(****************************************************************************************************<br>
© Syntegon Group.<br>
All rights reserved, also regarding any disposal, exploitation, reproduction, editing, distribution,<br>
as well as in the event of applications for industrial property rights.<br>
*****************************************************************************************************<br>
DESCRIPTION:<br>
Base of every robot (Delta, XTS gantry, XTS loop, Cartesian): zones plus the gripper fingers, m_SetFinger,<br>
m_SetFingerOffset (a finger's place on the flange) and m_ClearFingers, the limit area, m_SetLimitArea and<br>
m_ClearLimitArea, and the TCP limit area, m_SetTcpLimitArea and m_ClearTcpLimitArea. A derived FB tells where<br>
its fingers and its boxes lie through m_Fingers and m_LimitArea; an XTS loop has neither box.<br>
Not used directly.<br>
*****************************************************************************************************<br>
VERSION         ¦ DATE       ¦ NAME      ¦ CHANGE<br>
Syn_Visu 4.0.0  ¦ 2026-11-01 ¦ J.Willner ¦ New: fingers shared by all robots<br>
Syn_Visu 9.3.0  ¦ 2026-11-07 ¦ J.Willner ¦ Limit area shared by Delta, XTS gantry and Cartesian (was Delta only)<br>
Syn_Visu 9.4.0  ¦ 2026-11-09 ¦ J.Willner ¦ TCP limit area: m_SetTcpLimitArea, m_ClearTcpLimitArea<br>
Syn_Visu 9.4.1  ¦ 2026-11-09 ¦ J.Willner ¦ Limit area compares ignore padding: no config change from unchanged values<br>
Syn_Visu 9.5.0  ¦ 2026-11-11 ¦ J.Willner ¦ m_SetFingerOffset: a finger's place on the flange (ADR 0018)<br>
****************************************************************************************************)
FUNCTION_BLOCK ABSTRACT _FB_VisuRobot EXTENDS _FB_VisuZoneComponent

(****************************************************************************************************<br>
© Syntegon Group.<br>
All rights reserved, also regarding any disposal, exploitation, reproduction, editing, distribution,<br>
as well as in the event of applications for industrial property rights.<br>
*****************************************************************************************************<br>
DESCRIPTION:<br>
Removes the gripper definition. TRUE if there was one.<br>
****************************************************************************************************)
METHOD m_ClearFingers : BOOL
VAR
	p_TempCount							: POINTER TO UINT;
	p_TempFingers						: POINTER TO ARRAY[0..VISU_GlobalConst_Param.VISU_un_MAX_FINGERS - 1] OF ST_VisuFinger;
	TempEmpty							: ST_VisuFinger;
	un_TempIndex						: UINT;
END_VAR
m_ClearFingers := FALSE;
m_Fingers(vo_p_Count => p_TempCount, vo_p_Fingers => p_TempFingers);
IF p_TempCount = 0 OR p_TempFingers = 0 THEN
	RETURN;
END_IF
m_ClearFingers := p_TempCount^ > 0;
FOR un_TempIndex := 0 TO VISU_GlobalConst_Param.VISU_un_MAX_FINGERS - 1 DO
	p_TempFingers^[un_TempIndex] := TempEmpty;
END_FOR
p_TempCount^ := 0;
IF m_ClearFingers THEN
	m_NotifyConfigChanged();
END_IF
END_METHOD

(****************************************************************************************************<br>
© Syntegon Group.<br>
All rights reserved, also regarding any disposal, exploitation, reproduction, editing, distribution,<br>
as well as in the event of applications for industrial property rights.<br>
*****************************************************************************************************<br>
DESCRIPTION:<br>
Removes the limit area. TRUE if there was one.<br>
****************************************************************************************************)
METHOD m_ClearLimitArea : BOOL
VAR
	p_TempLimitArea						: POINTER TO ST_VisuLimitArea;
	TempEmpty							: ST_VisuLimitArea;
END_VAR
m_ClearLimitArea := FALSE;
m_LimitArea(vo_p_LimitArea => p_TempLimitArea);
IF p_TempLimitArea = 0 THEN
	RETURN;
END_IF
m_ClearLimitArea := p_TempLimitArea^.bActive;
(* Zeroed first: the MEMCMP below also compares the padding after bActive, which a method local leaves undefined. *)
Tc2_System.MEMSET(ADR(TempEmpty), 0, SIZEOF(TempEmpty));
IF Tc2_System.MEMCMP(ADR(TempEmpty), p_TempLimitArea, SIZEOF(TempEmpty)) <> 0 THEN
	p_TempLimitArea^ := TempEmpty;
	m_NotifyConfigChanged();
END_IF
END_METHOD

(****************************************************************************************************<br>
© Syntegon Group.<br>
All rights reserved, also regarding any disposal, exploitation, reproduction, editing, distribution,<br>
as well as in the event of applications for industrial property rights.<br>
*****************************************************************************************************<br>
DESCRIPTION:<br>
Removes the TCP limit area. TRUE if there was one.<br>
****************************************************************************************************)
METHOD m_ClearTcpLimitArea : BOOL
VAR
	p_TempTcpLimitArea					: POINTER TO ST_VisuLimitArea;
	TempEmpty							: ST_VisuLimitArea;
END_VAR
m_ClearTcpLimitArea := FALSE;
m_LimitArea(vo_p_TcpLimitArea => p_TempTcpLimitArea);
IF p_TempTcpLimitArea = 0 THEN
	RETURN;
END_IF
m_ClearTcpLimitArea := p_TempTcpLimitArea^.bActive;
(* Zeroed first: the MEMCMP below also compares the padding after bActive, which a method local leaves undefined. *)
Tc2_System.MEMSET(ADR(TempEmpty), 0, SIZEOF(TempEmpty));
IF Tc2_System.MEMCMP(ADR(TempEmpty), p_TempTcpLimitArea, SIZEOF(TempEmpty)) <> 0 THEN
	p_TempTcpLimitArea^ := TempEmpty;
	m_NotifyConfigChanged();
END_IF
END_METHOD

(****************************************************************************************************<br>
© Syntegon Group.<br>
All rights reserved, also regarding any disposal, exploitation, reproduction, editing, distribution,<br>
as well as in the event of applications for industrial property rights.<br>
*****************************************************************************************************<br>
DESCRIPTION:<br>
Where the gripper fingers lie in the derived FB's contract structure: vo_p_Count points to its<br>
nFingerCount, vo_p_Fingers to its aFingers.<br>
****************************************************************************************************)
METHOD PROTECTED ABSTRACT m_Fingers : BOOL
VAR_OUTPUT
	vo_p_Count							: POINTER TO UINT;
	vo_p_Fingers						: POINTER TO ARRAY[0..VISU_GlobalConst_Param.VISU_un_MAX_FINGERS - 1] OF ST_VisuFinger;
END_VAR
END_METHOD

(****************************************************************************************************<br>
© Syntegon Group.<br>
All rights reserved, also regarding any disposal, exploitation, reproduction, editing, distribution,<br>
as well as in the event of applications for industrial property rights.<br>
*****************************************************************************************************<br>
DESCRIPTION:<br>
Where the limit area and the TCP limit area lie in the derived FB's contract structure: vo_p_LimitArea points<br>
to its stLimitArea, vo_p_TcpLimitArea to its stTcpLimitArea; both are 0 for a robot without them (XTS loop: it<br>
has no working area of its own).<br>
****************************************************************************************************)
METHOD PROTECTED ABSTRACT m_LimitArea : BOOL
VAR_OUTPUT
	vo_p_LimitArea						: POINTER TO ST_VisuLimitArea;
	vo_p_TcpLimitArea					: POINTER TO ST_VisuLimitArea;
END_VAR
END_METHOD

(****************************************************************************************************<br>
© Syntegon Group.<br>
All rights reserved, also regarding any disposal, exploitation, reproduction, editing, distribution,<br>
as well as in the event of applications for industrial property rights.<br>
*****************************************************************************************************<br>
DESCRIPTION:<br>
Defines gripper finger vi_un_Finger (1-based): a cylinder hanging from the finger's pose along its local -Z.<br>
For XTS kinematics it is a finger of every mover's gripper. The finger count grows to vi_un_Finger.<br>
Its place on the gripper flange comes from m_SetFingerOffset and is kept here.<br>
*****************************************************************************************************<br>
OUTPUT VALUES:<br>
FALSE outside 1..VISU_GlobalConst_Param.VISU_un_MAX_FINGERS.<br>
****************************************************************************************************)
METHOD m_SetFinger : BOOL
VAR_INPUT
	vi_un_Finger						: UINT;	// [-] 1-based, as a product's nFingerId
	vi_lr_Diameter						: LREAL;	// [mm]
	vi_lr_Height						: LREAL;	// [mm] along the finger's local -Z
END_VAR
VAR
	p_TempCount							: POINTER TO UINT;
	p_TempFingers						: POINTER TO ARRAY[0..VISU_GlobalConst_Param.VISU_un_MAX_FINGERS - 1] OF ST_VisuFinger;
	TempFinger							: ST_VisuFinger;
END_VAR
m_SetFinger := FALSE;
IF vi_un_Finger = 0 OR vi_un_Finger > VISU_GlobalConst_Param.VISU_un_MAX_FINGERS THEN
	RETURN;
END_IF
m_Fingers(vo_p_Count => p_TempCount, vo_p_Fingers => p_TempFingers);
IF p_TempCount = 0 OR p_TempFingers = 0 THEN
	RETURN;
END_IF
TempFinger.fDiameter := vi_lr_Diameter;
TempFinger.fHeight := vi_lr_Height;
(* The offset stays as m_SetFingerOffset set it. *)
TempFinger.stOffset := p_TempFingers^[vi_un_Finger - 1].stOffset;
IF vi_un_Finger > p_TempCount^
OR Tc2_System.MEMCMP(ADR(TempFinger), ADR(p_TempFingers^[vi_un_Finger - 1]), SIZEOF(TempFinger)) <> 0
THEN
	p_TempFingers^[vi_un_Finger - 1] := TempFinger;
	p_TempCount^ := MAX(p_TempCount^, vi_un_Finger);
	m_NotifyConfigChanged();
END_IF
m_SetFinger := TRUE;
END_METHOD

(****************************************************************************************************<br>
© Syntegon Group.<br>
All rights reserved, also regarding any disposal, exploitation, reproduction, editing, distribution,<br>
as well as in the event of applications for industrial property rights.<br>
*****************************************************************************************************<br>
DESCRIPTION:<br>
Places finger vi_un_Finger (1-based, defined with m_SetFinger) on the gripper flange (ADR 0018): the position<br>
of its frame in the flange frame and its rotation about the flange's Z. The flange frame's -Z points to the<br>
product: a Delta's lies at the TCP with the robot's axes, a Cartesian robot's has the robot's axes, an XTS mover's<br>
turns with the mover. While the application reports no pose for the finger (m_SetFingerState, or an XTS track<br>
with m_SetFingersOnFlange), the visualisation draws it there. The config version only changes when a value does.<br>
*****************************************************************************************************<br>
OUTPUT VALUES:<br>
FALSE for a finger outside 1..the finger count.<br>
****************************************************************************************************)
METHOD m_SetFingerOffset : BOOL
VAR_INPUT
	vi_un_Finger						: UINT;	// [-] 1-based
	vi_lr_X								: LREAL;	// [mm] along the flange's X
	vi_lr_Y								: LREAL;	// [mm] along the flange's Y
	vi_lr_Z								: LREAL;	// [mm] along the flange's Z (towards the product: negative)
	vi_lr_Rz							: LREAL;	// [deg] about the flange's Z
END_VAR
VAR
	p_TempCount							: POINTER TO UINT;
	p_TempFingers						: POINTER TO ARRAY[0..VISU_GlobalConst_Param.VISU_un_MAX_FINGERS - 1] OF ST_VisuFinger;
	TempOffset							: ST_VisuPlanarPose;
END_VAR
m_SetFingerOffset := FALSE;
m_Fingers(vo_p_Count => p_TempCount, vo_p_Fingers => p_TempFingers);
IF p_TempCount = 0 OR p_TempFingers = 0 THEN
	RETURN;
END_IF
IF vi_un_Finger = 0 OR vi_un_Finger > p_TempCount^ THEN
	RETURN;
END_IF
TempOffset.fX := vi_lr_X;
TempOffset.fY := vi_lr_Y;
TempOffset.fZ := vi_lr_Z;
TempOffset.fRz := vi_lr_Rz;
IF Tc2_System.MEMCMP(ADR(TempOffset), ADR(p_TempFingers^[vi_un_Finger - 1].stOffset), SIZEOF(TempOffset)) <> 0 THEN
	p_TempFingers^[vi_un_Finger - 1].stOffset := TempOffset;
	m_NotifyConfigChanged();
END_IF
m_SetFingerOffset := TRUE;
END_METHOD

(****************************************************************************************************<br>
© Syntegon Group.<br>
All rights reserved, also regarding any disposal, exploitation, reproduction, editing, distribution,<br>
as well as in the event of applications for industrial property rights.<br>
*****************************************************************************************************<br>
DESCRIPTION:<br>
Sets and activates the limit area: an axis-aligned box in the robot frame (relative to its pose, the frame its<br>
working area is given in) that further restricts the working area. Delta, XTS gantry and Cartesian robot;<br>
an XTS loop has none. Equal bounds make a flat box. The config version only changes when a value does.<br>
*****************************************************************************************************<br>
OUTPUT VALUES:<br>
TRUE if anything changed; FALSE for a robot without a limit area (XTS loop).<br>
****************************************************************************************************)
METHOD m_SetLimitArea : BOOL
VAR_INPUT
	vi_lr_XMin							: LREAL;	// [mm] in the robot frame
	vi_lr_XMax							: LREAL;	// [mm]
	vi_lr_YMin							: LREAL;	// [mm]
	vi_lr_YMax							: LREAL;	// [mm]
	vi_lr_ZMin							: LREAL;	// [mm] relative to the pose (below it: negative)
	vi_lr_ZMax							: LREAL;	// [mm]
END_VAR
VAR
	p_TempLimitArea						: POINTER TO ST_VisuLimitArea;
	TempLimitArea						: ST_VisuLimitArea;
END_VAR
m_SetLimitArea := FALSE;
m_LimitArea(vo_p_LimitArea => p_TempLimitArea);
IF p_TempLimitArea = 0 THEN
	RETURN;
END_IF
(* Zeroed first: the MEMCMP below also compares the padding after bActive, which a method local leaves undefined. *)
Tc2_System.MEMSET(ADR(TempLimitArea), 0, SIZEOF(TempLimitArea));
TempLimitArea.fXMin := vi_lr_XMin;
TempLimitArea.fXMax := vi_lr_XMax;
TempLimitArea.fYMin := vi_lr_YMin;
TempLimitArea.fYMax := vi_lr_YMax;
TempLimitArea.fZMin := vi_lr_ZMin;
TempLimitArea.fZMax := vi_lr_ZMax;
TempLimitArea.bActive := TRUE;
IF Tc2_System.MEMCMP(ADR(TempLimitArea), p_TempLimitArea, SIZEOF(TempLimitArea)) <> 0 THEN
	p_TempLimitArea^ := TempLimitArea;
	m_NotifyConfigChanged();
	m_SetLimitArea := TRUE;
END_IF
END_METHOD

(****************************************************************************************************<br>
© Syntegon Group.<br>
All rights reserved, also regarding any disposal, exploitation, reproduction, editing, distribution,<br>
as well as in the event of applications for industrial property rights.<br>
*****************************************************************************************************<br>
DESCRIPTION:<br>
Sets and activates the TCP limit area: an axis-aligned box around the TCP (XTS gantry: around every mover's<br>
gripper flange), its bounds relative to the TCP along the axes of the robot frame. It moves with the TCP and<br>
never turns. The visualisation lights it up red with a message when it overlaps another robot's limit area or<br>
TCP limit area (also another mover's of the same gantry), or leaves the robot's own limit area. Delta, XTS<br>
gantry and Cartesian robot; an XTS loop has none. Equal bounds make a flat box. The config version only<br>
changes when a value does.<br>
*****************************************************************************************************<br>
OUTPUT VALUES:<br>
TRUE if anything changed; FALSE for a robot without a TCP limit area (XTS loop).<br>
****************************************************************************************************)
METHOD m_SetTcpLimitArea : BOOL
VAR_INPUT
	vi_lr_XMin							: LREAL;	// [mm] relative to the TCP, along the robot frame's X
	vi_lr_XMax							: LREAL;	// [mm]
	vi_lr_YMin							: LREAL;	// [mm]
	vi_lr_YMax							: LREAL;	// [mm]
	vi_lr_ZMin							: LREAL;	// [mm] relative to the TCP (below it: negative)
	vi_lr_ZMax							: LREAL;	// [mm]
END_VAR
VAR
	p_TempTcpLimitArea					: POINTER TO ST_VisuLimitArea;
	TempTcpLimitArea					: ST_VisuLimitArea;
END_VAR
m_SetTcpLimitArea := FALSE;
m_LimitArea(vo_p_TcpLimitArea => p_TempTcpLimitArea);
IF p_TempTcpLimitArea = 0 THEN
	RETURN;
END_IF
(* Zeroed first: the MEMCMP below also compares the padding after bActive, which a method local leaves undefined. *)
Tc2_System.MEMSET(ADR(TempTcpLimitArea), 0, SIZEOF(TempTcpLimitArea));
TempTcpLimitArea.fXMin := vi_lr_XMin;
TempTcpLimitArea.fXMax := vi_lr_XMax;
TempTcpLimitArea.fYMin := vi_lr_YMin;
TempTcpLimitArea.fYMax := vi_lr_YMax;
TempTcpLimitArea.fZMin := vi_lr_ZMin;
TempTcpLimitArea.fZMax := vi_lr_ZMax;
TempTcpLimitArea.bActive := TRUE;
IF Tc2_System.MEMCMP(ADR(TempTcpLimitArea), p_TempTcpLimitArea, SIZEOF(TempTcpLimitArea)) <> 0 THEN
	p_TempTcpLimitArea^ := TempTcpLimitArea;
	m_NotifyConfigChanged();
	m_SetTcpLimitArea := TRUE;
END_IF
END_METHOD

END_FUNCTION_BLOCK

(* stored: Version 1.1.0.1, ProductVersion 3.1.4026.18
   POU _FB_VisuRobot: Id {5ceb582b-104f-47cb-91fd-61b1cc207460}, SpecialFunc None
   Method m_ClearFingers: Id {c59c54bb-9b8a-4354-8e47-b266be81a7d2}
   Method m_ClearLimitArea: Id {860a5579-9f26-458c-b290-d105a32d5cba}
   Method m_ClearTcpLimitArea: Id {8f8cd439-d9ce-4c1d-b91b-58af4e37550c}
   Method m_Fingers: Id {a244e015-94d6-456e-b723-254a871e0b47}
   Method m_LimitArea: Id {422ae902-a026-4b53-81df-e5504829a257}
   Method m_SetFinger: Id {e7ffdbfc-b2ac-4437-abcd-43e830fe868a}
   Method m_SetFingerOffset: Id {fbf85459-e4a9-4ec0-bbc3-bc060bba20c4}
   Method m_SetLimitArea: Id {c83e3c90-d747-4568-a7bd-6b20d6038e33}
   Method m_SetTcpLimitArea: Id {3a6e8120-3b40-4865-afd0-0494858b88ec} *)
